   IF #Startup THEN
       "StationA".Access.Policy.Required[11] := 3;
       "StationB".Access.Policy.Required[11] := 3;
   END_IF;
   IF #Startup THEN
       IF NOT "FRK_AccessStorage".UsersCommissioned AND "FRK_LocalUsers".SchemaVersion = 0 AND "FRK_LocalUsers".Generation = 0 AND "FRK_LocalUsers".Checksum = DWORD#0 THEN
           "F_AccessBenchProvision"();
       END_IF;
       "StationA".Access.Policy.Required[2] := 1;
       "StationA".Access.Policy.Required[4] := 1;
       "StationA".Access.Policy.Required[5] := 1;
       "StationA".Access.Policy.Required[8] := 4;
       "StationA".Access.Policy.SessionTimeout := T#0ms;
       "StationB".Access.Policy.Required[2] := 1;
       "StationB".Access.Policy.Required[4] := 1;
       "StationB".Access.Policy.Required[5] := 1;
       "StationB".Access.Policy.Required[8] := 4;
       "StationB".Access.Policy.SessionTimeout := T#0ms;
       "GDB_AccessTest".HashData[0] := BYTE#16#00;
       "GDB_AccessTest".HashData[1] := BYTE#16#01;
       "GDB_AccessTest".HashData[2] := BYTE#16#02;
       "GDB_AccessTest".HashData[3] := BYTE#16#03;
       "GDB_AccessTest".HashData[4] := BYTE#16#04;
       "GDB_AccessTest".HashData[5] := BYTE#16#05;
       "GDB_AccessTest".HashData[6] := BYTE#16#06;
       "GDB_AccessTest".HashData[7] := BYTE#16#07;
       "GDB_AccessTest".HashData[8] := BYTE#16#08;
       "GDB_AccessTest".HashData[9] := BYTE#16#09;
       "GDB_AccessTest".HashData[10] := BYTE#16#0A;
       "GDB_AccessTest".HashData[11] := BYTE#16#0B;
       "GDB_AccessTest".HashData[12] := BYTE#16#0C;
       "GDB_AccessTest".HashData[13] := BYTE#16#0D;
       "GDB_AccessTest".HashData[14] := BYTE#16#0E;
       "GDB_AccessTest".HashData[15] := BYTE#16#0F;
       "GDB_AccessTest".HashData[16] := BYTE#16#10;
       "GDB_AccessTest".HashData[17] := BYTE#16#11;
       "GDB_AccessTest".HashData[18] := BYTE#16#12;
       "GDB_AccessTest".HashData[19] := BYTE#16#13;
       "GDB_AccessTest".HashData[20] := BYTE#16#14;
       "GDB_AccessTest".HashData[21] := BYTE#16#15;
       "GDB_AccessTest".HashData[22] := BYTE#16#16;
       "GDB_AccessTest".HashData[23] := BYTE#16#17;
       "GDB_AccessTest".HashData[24] := BYTE#16#18;
       "GDB_AccessTest".HashData[25] := BYTE#16#19;
       "GDB_AccessTest".HashData[26] := BYTE#16#1A;
       "GDB_AccessTest".HashData[27] := BYTE#16#1B;
       "GDB_AccessTest".HashData[28] := BYTE#16#1C;
       "GDB_AccessTest".HashData[29] := BYTE#16#1D;
       "GDB_AccessTest".HashData[30] := BYTE#16#1E;
       "GDB_AccessTest".HashData[31] := BYTE#16#1F;
       "GDB_AccessTest".HashData[32] := BYTE#16#20;
       "GDB_AccessTest".HashData[33] := BYTE#16#21;
       "GDB_AccessTest".HashData[34] := BYTE#16#22;
       "GDB_AccessTest".HashData[35] := BYTE#16#23;
       "GDB_AccessTest".HashData[36] := BYTE#16#24;
       "GDB_AccessTest".HashData[37] := BYTE#16#25;
       "GDB_AccessTest".HashData[38] := BYTE#16#26;
       "GDB_AccessTest".HashData[39] := BYTE#16#27;
       "GDB_AccessTest".HashData[40] := BYTE#16#28;
       "GDB_AccessTest".HashData[41] := BYTE#16#29;
       "GDB_AccessTest".HashData[42] := BYTE#16#2A;
       "GDB_AccessTest".HashData[43] := BYTE#16#2B;
       "GDB_AccessTest".HashData[44] := BYTE#16#2C;
       "GDB_AccessTest".HashData[45] := BYTE#16#2D;
       "GDB_AccessTest".HashData[46] := BYTE#16#2E;
       "GDB_AccessTest".HashData[47] := BYTE#16#2F;
       "GDB_AccessTest".HashOk := "FRK_Sha256Pin"(Data := "GDB_AccessTest".HashData, Size := 0, Digest := "GDB_AccessTest".Hash0);
       "GDB_AccessTest".HashData[0] := BYTE#16#61;
       "GDB_AccessTest".HashData[1] := BYTE#16#62;
       "GDB_AccessTest".HashData[2] := BYTE#16#63;
       "GDB_AccessTest".HashData[3] := BYTE#16#00;
       "GDB_AccessTest".HashData[4] := BYTE#16#00;
       "GDB_AccessTest".HashData[5] := BYTE#16#00;
       "GDB_AccessTest".HashData[6] := BYTE#16#00;
       "GDB_AccessTest".HashData[7] := BYTE#16#00;
       "GDB_AccessTest".HashData[8] := BYTE#16#00;
       "GDB_AccessTest".HashData[9] := BYTE#16#00;
       "GDB_AccessTest".HashData[10] := BYTE#16#00;
       "GDB_AccessTest".HashData[11] := BYTE#16#00;
       "GDB_AccessTest".HashData[12] := BYTE#16#00;
       "GDB_AccessTest".HashData[13] := BYTE#16#00;
       "GDB_AccessTest".HashData[14] := BYTE#16#00;
       "GDB_AccessTest".HashData[15] := BYTE#16#00;
       "GDB_AccessTest".HashData[16] := BYTE#16#00;
       "GDB_AccessTest".HashData[17] := BYTE#16#00;
       "GDB_AccessTest".HashData[18] := BYTE#16#00;
       "GDB_AccessTest".HashData[19] := BYTE#16#00;
       "GDB_AccessTest".HashData[20] := BYTE#16#00;
       "GDB_AccessTest".HashData[21] := BYTE#16#00;
       "GDB_AccessTest".HashData[22] := BYTE#16#00;
       "GDB_AccessTest".HashData[23] := BYTE#16#00;
       "GDB_AccessTest".HashData[24] := BYTE#16#00;
       "GDB_AccessTest".HashData[25] := BYTE#16#00;
       "GDB_AccessTest".HashData[26] := BYTE#16#00;
       "GDB_AccessTest".HashData[27] := BYTE#16#00;
       "GDB_AccessTest".HashData[28] := BYTE#16#00;
       "GDB_AccessTest".HashData[29] := BYTE#16#00;
       "GDB_AccessTest".HashData[30] := BYTE#16#00;
       "GDB_AccessTest".HashData[31] := BYTE#16#00;
       "GDB_AccessTest".HashData[32] := BYTE#16#00;
       "GDB_AccessTest".HashData[33] := BYTE#16#00;
       "GDB_AccessTest".HashData[34] := BYTE#16#00;
       "GDB_AccessTest".HashData[35] := BYTE#16#00;
       "GDB_AccessTest".HashData[36] := BYTE#16#00;
       "GDB_AccessTest".HashData[37] := BYTE#16#00;
       "GDB_AccessTest".HashData[38] := BYTE#16#00;
       "GDB_AccessTest".HashData[39] := BYTE#16#00;
       "GDB_AccessTest".HashData[40] := BYTE#16#00;
       "GDB_AccessTest".HashData[41] := BYTE#16#00;
       "GDB_AccessTest".HashData[42] := BYTE#16#00;
       "GDB_AccessTest".HashData[43] := BYTE#16#00;
       "GDB_AccessTest".HashData[44] := BYTE#16#00;
       "GDB_AccessTest".HashData[45] := BYTE#16#00;
       "GDB_AccessTest".HashData[46] := BYTE#16#00;
       "GDB_AccessTest".HashData[47] := BYTE#16#00;
       "GDB_AccessTest".HashOk := "FRK_Sha256Pin"(Data := "GDB_AccessTest".HashData, Size := 3, Digest := "GDB_AccessTest".Hash1);
       "GDB_AccessTest".HashData[0] := BYTE#16#00;
       "GDB_AccessTest".HashData[1] := BYTE#16#01;
       "GDB_AccessTest".HashData[2] := BYTE#16#02;
       "GDB_AccessTest".HashData[3] := BYTE#16#03;
       "GDB_AccessTest".HashData[4] := BYTE#16#04;
       "GDB_AccessTest".HashData[5] := BYTE#16#05;
       "GDB_AccessTest".HashData[6] := BYTE#16#06;
       "GDB_AccessTest".HashData[7] := BYTE#16#07;
       "GDB_AccessTest".HashData[8] := BYTE#16#08;
       "GDB_AccessTest".HashData[9] := BYTE#16#09;
       "GDB_AccessTest".HashData[10] := BYTE#16#0A;
       "GDB_AccessTest".HashData[11] := BYTE#16#0B;
       "GDB_AccessTest".HashData[12] := BYTE#16#0C;
       "GDB_AccessTest".HashData[13] := BYTE#16#0D;
       "GDB_AccessTest".HashData[14] := BYTE#16#0E;
       "GDB_AccessTest".HashData[15] := BYTE#16#0F;
       "GDB_AccessTest".HashData[16] := BYTE#16#10;
       "GDB_AccessTest".HashData[17] := BYTE#16#11;
       "GDB_AccessTest".HashData[18] := BYTE#16#12;
       "GDB_AccessTest".HashData[19] := BYTE#16#13;
       "GDB_AccessTest".HashData[20] := BYTE#16#14;
       "GDB_AccessTest".HashData[21] := BYTE#16#15;
       "GDB_AccessTest".HashData[22] := BYTE#16#16;
       "GDB_AccessTest".HashData[23] := BYTE#16#17;
       "GDB_AccessTest".HashData[24] := BYTE#16#18;
       "GDB_AccessTest".HashData[25] := BYTE#16#19;
       "GDB_AccessTest".HashData[26] := BYTE#16#1A;
       "GDB_AccessTest".HashData[27] := BYTE#16#1B;
       "GDB_AccessTest".HashData[28] := BYTE#16#1C;
       "GDB_AccessTest".HashData[29] := BYTE#16#1D;
       "GDB_AccessTest".HashData[30] := BYTE#16#1E;
       "GDB_AccessTest".HashData[31] := BYTE#16#1F;
       "GDB_AccessTest".HashData[32] := BYTE#16#20;
       "GDB_AccessTest".HashData[33] := BYTE#16#21;
       "GDB_AccessTest".HashData[34] := BYTE#16#22;
       "GDB_AccessTest".HashData[35] := BYTE#16#23;
       "GDB_AccessTest".HashData[36] := BYTE#16#24;
       "GDB_AccessTest".HashData[37] := BYTE#16#25;
       "GDB_AccessTest".HashData[38] := BYTE#16#26;
       "GDB_AccessTest".HashData[39] := BYTE#16#27;
       "GDB_AccessTest".HashData[40] := BYTE#16#28;
       "GDB_AccessTest".HashData[41] := BYTE#16#29;
       "GDB_AccessTest".HashData[42] := BYTE#16#2A;
       "GDB_AccessTest".HashData[43] := BYTE#16#2B;
       "GDB_AccessTest".HashData[44] := BYTE#16#2C;
       "GDB_AccessTest".HashData[45] := BYTE#16#2D;
       "GDB_AccessTest".HashData[46] := BYTE#16#2E;
       "GDB_AccessTest".HashData[47] := BYTE#16#2F;
       "GDB_AccessTest".HashOk := "FRK_Sha256Pin"(Data := "GDB_AccessTest".HashData, Size := 32, Digest := "GDB_AccessTest".Hash2);
       "GDB_AccessTest".HashData[0] := BYTE#16#00;
       "GDB_AccessTest".HashData[1] := BYTE#16#01;
       "GDB_AccessTest".HashData[2] := BYTE#16#02;
       "GDB_AccessTest".HashData[3] := BYTE#16#03;
       "GDB_AccessTest".HashData[4] := BYTE#16#04;
       "GDB_AccessTest".HashData[5] := BYTE#16#05;
       "GDB_AccessTest".HashData[6] := BYTE#16#06;
       "GDB_AccessTest".HashData[7] := BYTE#16#07;
       "GDB_AccessTest".HashData[8] := BYTE#16#08;
       "GDB_AccessTest".HashData[9] := BYTE#16#09;
       "GDB_AccessTest".HashData[10] := BYTE#16#0A;
       "GDB_AccessTest".HashData[11] := BYTE#16#0B;
       "GDB_AccessTest".HashData[12] := BYTE#16#0C;
       "GDB_AccessTest".HashData[13] := BYTE#16#0D;
       "GDB_AccessTest".HashData[14] := BYTE#16#0E;
       "GDB_AccessTest".HashData[15] := BYTE#16#0F;
       "GDB_AccessTest".HashData[16] := BYTE#16#10;
       "GDB_AccessTest".HashData[17] := BYTE#16#11;
       "GDB_AccessTest".HashData[18] := BYTE#16#12;
       "GDB_AccessTest".HashData[19] := BYTE#16#13;
       "GDB_AccessTest".HashData[20] := BYTE#16#14;
       "GDB_AccessTest".HashData[21] := BYTE#16#15;
       "GDB_AccessTest".HashData[22] := BYTE#16#16;
       "GDB_AccessTest".HashData[23] := BYTE#16#17;
       "GDB_AccessTest".HashData[24] := BYTE#16#18;
       "GDB_AccessTest".HashData[25] := BYTE#16#19;
       "GDB_AccessTest".HashData[26] := BYTE#16#1A;
       "GDB_AccessTest".HashData[27] := BYTE#16#1B;
       "GDB_AccessTest".HashData[28] := BYTE#16#1C;
       "GDB_AccessTest".HashData[29] := BYTE#16#1D;
       "GDB_AccessTest".HashData[30] := BYTE#16#1E;
       "GDB_AccessTest".HashData[31] := BYTE#16#1F;
       "GDB_AccessTest".HashData[32] := BYTE#16#20;
       "GDB_AccessTest".HashData[33] := BYTE#16#21;
       "GDB_AccessTest".HashData[34] := BYTE#16#22;
       "GDB_AccessTest".HashData[35] := BYTE#16#23;
       "GDB_AccessTest".HashData[36] := BYTE#16#24;
       "GDB_AccessTest".HashData[37] := BYTE#16#25;
       "GDB_AccessTest".HashData[38] := BYTE#16#26;
       "GDB_AccessTest".HashData[39] := BYTE#16#27;
       "GDB_AccessTest".HashData[40] := BYTE#16#28;
       "GDB_AccessTest".HashData[41] := BYTE#16#29;
       "GDB_AccessTest".HashData[42] := BYTE#16#2A;
       "GDB_AccessTest".HashData[43] := BYTE#16#2B;
       "GDB_AccessTest".HashData[44] := BYTE#16#2C;
       "GDB_AccessTest".HashData[45] := BYTE#16#2D;
       "GDB_AccessTest".HashData[46] := BYTE#16#2E;
       "GDB_AccessTest".HashData[47] := BYTE#16#2F;
       "GDB_AccessTest".HashOk := "FRK_Sha256Pin"(Data := "GDB_AccessTest".HashData, Size := 48, Digest := "GDB_AccessTest".Hash3);
       "GDB_RoutingTest".PermitOne := TRUE;
       "GDB_RoutingTest".PermitTwo := TRUE;
       "GDB_RoutingTest".RootManualPermit := TRUE;
       "GDB_RoutingTest".NestedFinish := FALSE;
       "GDB_RoutingTest".InnerFinish := FALSE;
       "GDB_RoutingTest".NestedAccessLock := FALSE;
       #ResultCode := RD_SYS_T(OUT => #StartupStamp);
       IF #ResultCode = 0 THEN
           "GDB_UnitTest".BootStamp := DTL_TO_LDT(#StartupStamp);
       END_IF;
       "GDB_UnitTest".Restarts := "GDB_UnitTest".Restarts + 1;
       "GDB_UnitTest".FinishCycle := FALSE;
       "GDB_UnitTest".Permit := TRUE;
       "GDB_UnitTest".FaultRoot := FALSE;
       "GDB_UnitTest".ExitHold := FALSE;
       "GDB_UnitTest".IssueChild := FALSE;
       "GDB_UnitTest".LockStart := FALSE;
       "GDB_UnitTest".ChildCommand := 2;
       "GDB_UnitTest".Verdict := 1;
       "GDB_UnitTest".Reason := 2003;
       "GDB_UnitTest".CarrierControl := 0;
       "FRK_UnitSetLocalCarrier"(Unit := "StationA".Unit,
                                 Index := 1);
   END_IF;
   "GDB_FraktalHal".Data.StationA.Cell.Clamp.Finish := "GDB_UnitTest".FinishCycle;
   "GDB_FraktalHal".Data.StationA.Cell.Clamp.Permit := "GDB_UnitTest".Permit;
   "GDB_FraktalHal".Data.StationA.Cell.Clamp.ExitHold := "GDB_UnitTest".ExitHold;
   "GDB_FraktalHal".Data.StationA.Cell.Clamp.BackgroundFault := "GDB_UnitTest".FaultRoot;
   "GDB_FraktalHal".Data.StationA.Cell.Clamp.Verdict := "GDB_UnitTest".Verdict;
   "GDB_FraktalHal".Data.StationA.Cell.Clamp.Diag.ReasonCode := "GDB_UnitTest".Reason;
   "GDB_FraktalHal".Data.StationA.Cell.Clamp.Diag.Description := WSTRING#'test.start.permit';
   "GDB_FraktalHal".Data.StationA.Cell.Clamp.Diag.SourcePath := WSTRING#'StationA.Cell.Clamp';
   IF "GDB_UnitTest".IssueChild THEN
       "StationA".Cell.Clamp.Command := "GDB_UnitTest".ChildCommand;
       "StationA".Cell.Clamp.Execute := TRUE;
       "GDB_UnitTest".IssueChild := FALSE;
   END_IF;
   CASE "GDB_UnitTest".CarrierControl OF
       1:
           "FRK_UnitSetLocalCarrier"(Unit := "StationA".Unit,
                                     Index := 1);
       2:
           "FRK_Carriers".Slots[1].Enabled := FALSE;
       3:
           "FRK_Carriers".Slots[1].Context.Uid := 'other';
       ELSE
           "GDB_UnitTest".CarrierControl := 0;
   END_CASE;
   "GDB_UnitTest".CarrierControl := 0;
   "GDB_FraktalHal".Data.StationA.Cell.Gate.Permit := "GDB_RoutingTest".PermitOne;
   IF "GDB_RoutingTest".PermitTwo THEN
       "GDB_FraktalHal".Data.StationA.Cell.Gate.Sample := 0;
   ELSE
       "GDB_FraktalHal".Data.StationA.Cell.Gate.Sample := 1;
   END_IF;
   "GDB_FraktalHal".Data.StationA.Cell.Gate.Diag.ReasonCode := 2002;
   "GDB_FraktalHal".Data.StationA.Cell.Gate.Diag.Description := WSTRING#'test.manual.first';
   "GDB_FraktalHal".Data.StationA.Cell.Gate.LaterDiag.ReasonCode := 2003;
   "GDB_FraktalHal".Data.StationA.Cell.Gate.LaterDiag.Description := WSTRING#'test.manual.second';
   "GDB_FraktalHal".Data.StationA.Satellite.Cell.Clamp.Permit := "GDB_RoutingTest".RootManualPermit;
   "GDB_FraktalHal".Data.StationA.Satellite.Cell.Clamp.Diag.SourcePath := WSTRING#'StationA.Satellite.Cell.Clamp';
   "GDB_FraktalHal".Data.StationA.Satellite.Cell.Clamp.Diag.Description := WSTRING#'test.nested.permit';
   "GDB_FraktalHal".Data.StationA.Satellite.Cell.Clamp.Diag.ReasonCode := 2002;
   "GDB_FraktalHal".Data.StationA.Satellite.Inner.Cell.Clamp.Permit := TRUE;
   "GDB_FraktalHal".Data.StationA.Satellite.Cell.Clamp.Finish := "GDB_RoutingTest".NestedFinish;
   "GDB_FraktalHal".Data.StationA.Satellite.Inner.Cell.Clamp.Finish := "GDB_RoutingTest".InnerFinish;
   IF "GDB_RoutingTest".NestedAccessLock THEN
       "StationA".Satellite.Access.Policy.Required[5] := 4;
   ELSE
       "StationA".Satellite.Access.Policy.Required[5] := 0;
   END_IF;
   IF "GDB_RoutingTest".LocalPulse THEN
       "GDB_RoutingTest".LocalRequest.Kind := "GDB_RoutingTest".LocalKind;
       "GDB_RoutingTest".LocalRequest.IntValue := "GDB_RoutingTest".LocalValue;
       "FRK_UnitOperation"(Core := "StationA".Satellite.Core,
                           Unit := "StationA".Satellite.Unit,
                           Status := "StationA".Satellite.Status,
                           Policy := "StationA".Satellite.ModePolicy,
                           Access := "StationA".Satellite.Access,
                           Supported := "StationA".Satellite.SupportedModesPublished,
                           Request := "GDB_RoutingTest".LocalRequest,
                           Response := "FRK_UnitScratch".Response,
                           Trusted := FALSE);
       "GDB_RoutingTest".LocalAccepted := "FRK_UnitScratch".Response.Accepted;
       "GDB_RoutingTest".LocalFirstKind := -1;
       IF "FRK_UnitScratch".Response.Report.Count > 0 THEN
           "GDB_RoutingTest".LocalFirstKind := "FRK_UnitScratch".Response.Report.Reasons[1].Kind;
       END_IF;
       "GDB_RoutingTest".LocalPulse := FALSE;
   END_IF;
   "StationA".Access.ProviderEnabled := NOT "GDB_AccessTest".ProviderOff;
   "StationB".Access.ProviderEnabled := NOT "GDB_AccessTest".ProviderOff;
   "StationA".AlarmLog.SinkEnabled := TRUE;
   "StationB".AlarmLog.SinkEnabled := TRUE;
   "GDB_FraktalHal".Data.StationA.Cell.Clamp.Sample := "GDB_StateAlarmTest".Position;
   IF "GDB_StateAlarmTest".ClearLog THEN
       "FRK_AlarmBegin"(AlarmLog := "StationA".AlarmLog,
                        Startup := TRUE);
       "GDB_StateAlarmTest".SinkCome := 0;
       "GDB_StateAlarmTest".SinkClose := 0;
       "GDB_StateAlarmTest".ClearLog := FALSE;
   END_IF;
   IF "GDB_StateAlarmTest".RaisePulse THEN
       "GDB_StateAlarmTest".Slot := "FRK_AlarmRaise"(AlarmLog := "StationA".AlarmLog, Diag := "GDB_StateAlarmTest".Diag, ResetClass := "GDB_StateAlarmTest".ResetClass);
       "GDB_StateAlarmTest".RaisePulse := FALSE;
   END_IF;
   IF "GDB_StateAlarmTest".GonePulse THEN
       "GDB_StateAlarmTest".GoneAccepted := "FRK_AlarmGone"(AlarmLog := "StationA".AlarmLog, Slot := "GDB_StateAlarmTest".Slot);
       "GDB_StateAlarmTest".GonePulse := FALSE;
   END_IF;
   IF "GDB_StateAlarmTest".FillPulse THEN
       FOR #SlotIndex := 1 TO "GDB_StateAlarmTest".FillCount DO
           #Taken := "FRK_AlarmRaise"(AlarmLog := "StationA".AlarmLog, Diag := "GDB_StateAlarmTest".Diag, ResetClass := "GDB_StateAlarmTest".ResetClass);
           IF "GDB_StateAlarmTest".ResetClass = 0 THEN
               #Accepted := "FRK_AlarmGone"(AlarmLog := "StationA".AlarmLog, Slot := #Taken);
           END_IF;
       END_FOR;
       "GDB_StateAlarmTest".FillPulse := FALSE;
   END_IF;
   IF "GDB_StateAlarmTest".CauseLive THEN
       IF "GDB_StateAlarmTest".CauseSlot = 0 THEN
           "GDB_StateAlarmTest".CauseSlot := "FRK_AlarmRaise"(AlarmLog := "StationA".AlarmLog, Diag := "GDB_StateAlarmTest".Diag, ResetClass := 1);
       ELSIF "StationA".AlarmLog.Active["GDB_StateAlarmTest".CauseSlot].State = 0 THEN
           "GDB_StateAlarmTest".CauseSlot := "FRK_AlarmRaise"(AlarmLog := "StationA".AlarmLog, Diag := "GDB_StateAlarmTest".Diag, ResetClass := 1);
       END_IF;
   ELSIF "GDB_StateAlarmTest".CauseSlot > 0 THEN
       #Accepted := "FRK_AlarmGone"(AlarmLog := "StationA".AlarmLog, Slot := "GDB_StateAlarmTest".CauseSlot);
       "GDB_StateAlarmTest".CauseSlot := 0;
   END_IF;
   "FRK_StateSweep"(Flags := "GDB_StateAlarmTest".StandaloneFlags,
                    Count := "GDB_StateAlarmTest".StandaloneCount,
                    Touched := "GDB_StateAlarmTest".Touched,
                    Startup := #Startup);
   IF "GDB_StateAlarmTest".PublishState THEN
       "GDB_StateAlarmTest".StandaloneReturn := "FRK_State"(Idx := "GDB_StateAlarmTest".StateIndex, Key := 'project.state.atHome', Ok := "GDB_StateAlarmTest".StateValue, Flags := "GDB_StateAlarmTest".StandaloneFlags, Count := "GDB_StateAlarmTest".StandaloneCount, Touched := "GDB_StateAlarmTest".Touched);
   END_IF;
   "FRK_ConfigRuntime".Unavailable := "GDB_ConfigTest".Unavailable;
   IF "GDB_ConfigTest".BlockRestore THEN
       "StationA".ConfigPersist.RestorePolicy := 1;
   ELSE
       "StationA".ConfigPersist.RestorePolicy := 0;
   END_IF;
   IF "GDB_ConfigTest".CorruptPulse THEN
       "GDB_ConfigTest".CorruptSlot := "FRK_ConfigFind"(Scope := "GDB_ConfigTest".CorruptScope, Key := "GDB_ConfigTest".CorruptKey, ModelCode := "GDB_ConfigTest".CorruptModel);
       IF "GDB_ConfigTest".CorruptSlot > 0 THEN
           "FRK_ConfigStore".Rows["GDB_ConfigTest".CorruptSlot].SchemaVersion := "GDB_ConfigTest".CorruptSchema;
           "FRK_ConfigStore".Rows["GDB_ConfigTest".CorruptSlot].Record.ValueText := "GDB_ConfigTest".CorruptText;
       END_IF;
       "GDB_ConfigTest".CorruptPulse := FALSE;
   END_IF;
END_FUNCTION

FUNCTION "F_ConfigSetBench" : Void   // FC173, SCL
{ S7_Optimized_Access := 'TRUE' }
VERSION : 0.1
// Test-only tampering: the production retained store stays inaccessible.
// stored: AutoNumber true, IsIECCheckEnabled false, SetENOAutomatically false, UDAEnableTagReadback false
   VAR_TEMP
      Slot : Int;
      Index : Int;
   END_VAR
BEGIN

   IF NOT "GDB_ConfigSetTest".Corrupt THEN
       RETURN;
   END_IF;
   "GDB_ConfigSetTest".Corrupt := FALSE;
   #Slot := "FRK_SetFind"(RootIndex := 1, SetName := "GDB_ConfigSetTest".SetName);
   "GDB_ConfigSetTest".Slot := #Slot;
   IF #Slot = 0 THEN
       RETURN;
   END_IF;
   #Index := "FRK_SetStore".Sets[1, #Slot].Info.RecordCount;
   "GDB_ConfigSetTest".RecordScope := "FRK_SetStore".Sets[1, #Slot].Records[#Index].Scope;
   "GDB_ConfigSetTest".RecordKey := "FRK_SetStore".Sets[1, #Slot].Records[#Index].WriteKey;
   CASE "GDB_ConfigSetTest".Field OF
       1:
           "FRK_SetStore".Sets[1, #Slot].Records[#Index].ValueText := "GDB_ConfigSetTest".Text;
       2:
           "FRK_SetStore".Sets[1, #Slot].Records[#Index].Revision := 99;
       3:
           "FRK_SetStore".Sets[1, #Slot].Records[#Index].ValueType := 99;
       4:
           "FRK_SetStore".Sets[1, #Slot].Records[#Index].WriteKey := 'unknown';
       5:
           "FRK_SetStore".Sets[1, #Slot].Records[#Index].Scope := 'StationB';
       6:
           "FRK_SetStore".Sets[1, #Slot].Info.RecordCount := #Index - 1;
       7:
           "FRK_SetStore".Sets[1, #Slot].Records[#Index] := "FRK_SetStore".Sets[1, #Slot].Records[1];
       ELSE
           RETURN;
   END_CASE;
END_FUNCTION

FUNCTION "F_DecisionBench" : Void   // FC172, SCL
{ S7_Optimized_Access := 'TRUE' }
VERSION : 0.1
// stored: AutoNumber true, IsIECCheckEnabled false, SetENOAutomatically false, UDAEnableTagReadback false
   VAR_TEMP
      Root : DInt;
      Peer : DInt;
      Nested : DInt;
      Slot : Int;
      CaseNo : Int;
      RootPath : WString[255];
      PeerPath : WString[255];
      NestedPath : WString[255];
      "A" : Bool;
      "B" : Bool;
      C : Bool;
      Ok : Bool;
      Answer : Int;
      Head : Int;
   END_VAR
BEGIN

   IF "GDB_DecisionTest".Done OR "FRK_Registry".Fault THEN
       RETURN;
   END_IF;
   #Root := "StationA".Core.RegIndex;
   #Peer := "StationB".Core.RegIndex;
   #Nested := "StationA".Satellite.Core.RegIndex;
   IF #Root <= 0 OR #Peer <= 0 OR #Nested <= 0 THEN
       RETURN;
   END_IF;
   #RootPath := STRING_TO_WSTRING("StationA".Status.Name);
   #PeerPath := STRING_TO_WSTRING("StationB".Status.Name);
   #NestedPath := STRING_TO_WSTRING("StationA".Satellite.Status.Name);
   #Slot := "FRK_DecisionRoot"(Owner := #Root, Create := TRUE);
   "GDB_DecisionTest".Total := 28;
   FOR #CaseNo := 1 TO 28 DO
       "FRK_DecisionCyclic"(Owner := #Root,
                            Busy := FALSE,
                            Reset := TRUE,
                            AlarmLog := "GDB_DecisionTest".Log);
       "FRK_DecisionCyclic"(Owner := #Peer,
                            Busy := FALSE,
                            Reset := TRUE,
                            AlarmLog := "GDB_DecisionTest".Log);
       "GDB_DecisionTest".WorkRequest := "FRK_Decisions".EmptyRequest;
       "GDB_DecisionTest".WorkRequest.Prompt := WSTRING#'test.decision.prompt';
       "GDB_DecisionTest".WorkRequest.Options[1] := 'test.decision.optionOne';
       "GDB_DecisionTest".WorkRequest.Options[2] := 'test.decision.optionTwo';
       "GDB_DecisionTest".WorkHmiRequest := "GDB_DecisionTest".EmptyHmiRequest;
       "GDB_DecisionTest".WorkHmiResponse := "GDB_DecisionTest".EmptyHmiResponse;
       "GDB_DecisionTest".WorkReport := "GDB_DecisionTest".EmptyReport;
       "GDB_DecisionTest".WorkPublished := "FRK_Decisions".EmptyRequest;
       "GDB_DecisionTest".WorkReport.Count := 0;
       "GDB_DecisionTest".WorkReport.Released := TRUE;
       #Ok := FALSE;
       CASE #CaseNo OF
           1: // invalid_owner
               #A := "FRK_DecisionAsk"(Owner := 0, OwnerPath := #RootPath, Request := "GDB_DecisionTest".WorkRequest, AlarmLog := "GDB_DecisionTest".Log);
               #Ok := NOT #A;
           2: // root_publication
               #A := "FRK_DecisionAsk"(Owner := #Root, OwnerPath := #RootPath, Request := "GDB_DecisionTest".WorkRequest, AlarmLog := "GDB_DecisionTest".Log);
               "FRK_DecisionPublish"(Owner := #Root,
                                     Decision := "GDB_DecisionTest".WorkPublished,
                                     DecisionAnswer := #Answer);
               #Ok := #A AND "GDB_DecisionTest".WorkPublished.Prompt = "GDB_DecisionTest".WorkRequest.Prompt AND "GDB_DecisionTest".WorkPublished.SourcePath = #RootPath AND #Answer = 0;
           3: // idempotent_no_flood
               #A := "FRK_DecisionAsk"(Owner := #Root, OwnerPath := #RootPath, Request := "GDB_DecisionTest".WorkRequest, AlarmLog := "GDB_DecisionTest".Log);
               #Head := "GDB_DecisionTest".Log.RingHead;
               #A := "FRK_DecisionAsk"(Owner := #Root, OwnerPath := #RootPath, Request := "GDB_DecisionTest".WorkRequest, AlarmLog := "GDB_DecisionTest".Log);
               #Ok := #A AND #Head = "GDB_DecisionTest".Log.RingHead;
           4: // overlap_preserves_first
               #A := "FRK_DecisionAsk"(Owner := #Root, OwnerPath := #RootPath, Request := "GDB_DecisionTest".WorkRequest, AlarmLog := "GDB_DecisionTest".Log);
               "GDB_DecisionTest".WorkRequest.Prompt := WSTRING#'test.decision.different';
               #A := "FRK_DecisionAsk"(Owner := #Root, OwnerPath := #RootPath, Request := "GDB_DecisionTest".WorkRequest, AlarmLog := "GDB_DecisionTest".Log);
               #Head := "GDB_DecisionTest".Log.RingHead;
               #B := #A;
               #A := "FRK_DecisionAsk"(Owner := #Root, OwnerPath := #RootPath, Request := "GDB_DecisionTest".WorkRequest, AlarmLog := "GDB_DecisionTest".Log);
               "FRK_DecisionPublish"(Owner := #Root,
                                     Decision := "GDB_DecisionTest".WorkPublished,
                                     DecisionAnswer := #Answer);
               #Ok := NOT #B AND NOT #A AND "GDB_DecisionTest".WorkPublished.Prompt = WSTRING#'test.decision.prompt' AND #Head = "GDB_DecisionTest".Log.RingHead;
           5: // nested_request_root_mirror
               #A := "FRK_DecisionAsk"(Owner := #Nested, OwnerPath := #NestedPath, Request := "GDB_DecisionTest".WorkRequest, AlarmLog := "GDB_DecisionTest".Log);
               "FRK_DecisionPublish"(Owner := #Root,
                                     Decision := "GDB_DecisionTest".WorkPublished,
                                     DecisionAnswer := #Answer);
               #B := "GDB_DecisionTest".WorkPublished.SourcePath = #NestedPath;
               "FRK_DecisionPublish"(Owner := #Nested,
                                     Decision := "GDB_DecisionTest".WorkPublished,
                                     DecisionAnswer := #Answer);
               #Ok := #A AND #B AND "GDB_DecisionTest".WorkPublished.Prompt = WSTRING#'';
           6: // peer_roots_independent
               #A := "FRK_DecisionAsk"(Owner := #Root, OwnerPath := #RootPath, Request := "GDB_DecisionTest".WorkRequest, AlarmLog := "GDB_DecisionTest".Log);
               "GDB_DecisionTest".WorkRequest.Prompt := WSTRING#'test.decision.peer';
               #B := "FRK_DecisionAsk"(Owner := #Peer, OwnerPath := #PeerPath, Request := "GDB_DecisionTest".WorkRequest, AlarmLog := "GDB_DecisionTest".Log);
               "FRK_DecisionPublish"(Owner := #Root,
                                     Decision := "GDB_DecisionTest".WorkPublished,
                                     DecisionAnswer := #Answer);
               #Ok := #A AND #B AND "GDB_DecisionTest".WorkPublished.Prompt = WSTRING#'test.decision.prompt';
               "FRK_DecisionPublish"(Owner := #Peer,
                                     Decision := "GDB_DecisionTest".WorkPublished,
                                     DecisionAnswer := #Answer);
               #Ok := #Ok AND "GDB_DecisionTest".WorkPublished.Prompt = WSTRING#'test.decision.peer';
           7: // zero_timeout_indefinite
               #A := "FRK_DecisionAsk"(Owner := #Root, OwnerPath := #RootPath, Request := "GDB_DecisionTest".WorkRequest, AlarmLog := "GDB_DecisionTest".Log);
               "FRK_Decisions".Slots[#Slot].AskedAt := "FRK_Clock".NowMs - 5000;
               "FRK_DecisionCyclic"(Owner := #Root,
                                    Busy := TRUE,
                                    Reset := FALSE,
                                    AlarmLog := "GDB_DecisionTest".Log);
               "FRK_DecisionPublish"(Owner := #Root,
                                     Decision := "GDB_DecisionTest".WorkPublished,
                                     DecisionAnswer := #Answer);
               #Ok := #A AND #Answer = 0 AND "GDB_DecisionTest".WorkPublished.Prompt <> WSTRING#'';
           8: // finite_timeout_default
               "GDB_DecisionTest".WorkRequest.Timeout := T#2ms;
               "GDB_DecisionTest".WorkRequest.Default := 2;
               #A := "FRK_DecisionAsk"(Owner := #Root, OwnerPath := #RootPath, Request := "GDB_DecisionTest".WorkRequest, AlarmLog := "GDB_DecisionTest".Log);
               "FRK_Decisions".Slots[#Slot].AskedAt := "FRK_Clock".NowMs - 5;
               "FRK_DecisionCyclic"(Owner := #Root,
                                    Busy := TRUE,
                                    Reset := FALSE,
                                    AlarmLog := "GDB_DecisionTest".Log);
               #Answer := "FRK_DecisionTake"(Owner := #Root, AlarmLog := "GDB_DecisionTest".Log);
               #Ok := #A AND #Answer = 2;
           9: // finite_requires_default
               "GDB_DecisionTest".WorkRequest.Timeout := T#2ms;
               #A := "FRK_DecisionAsk"(Owner := #Root, OwnerPath := #RootPath, Request := "GDB_DecisionTest".WorkRequest, AlarmLog := "GDB_DecisionTest".Log);
               #Ok := NOT #A;
           10: // default_must_be_offered
               "GDB_DecisionTest".WorkRequest.Default := 3;
               #A := "FRK_DecisionAsk"(Owner := #Root, OwnerPath := #RootPath, Request := "GDB_DecisionTest".WorkRequest, AlarmLog := "GDB_DecisionTest".Log);
               #Ok := NOT #A;
           11: // negative_timeout_rejected
               "GDB_DecisionTest".WorkRequest.Timeout := T#-1ms;
               #A := "FRK_DecisionAsk"(Owner := #Root, OwnerPath := #RootPath, Request := "GDB_DecisionTest".WorkRequest, AlarmLog := "GDB_DecisionTest".Log);
               #Ok := NOT #A;
           12: // option_zero_rejected
               #A := "FRK_DecisionAsk"(Owner := #Root, OwnerPath := #RootPath, Request := "GDB_DecisionTest".WorkRequest, AlarmLog := "GDB_DecisionTest".Log);
               "GDB_DecisionTest".WorkReport.Released := TRUE;
               #B := "FRK_DecisionSubmit"(Owner := #Root, OwnerPath := #RootPath, Option := 0, Busy := TRUE, Permit := TRUE, Report := "GDB_DecisionTest".WorkReport);
               #Ok := #A AND NOT #B AND NOT "GDB_DecisionTest".WorkReport.Released;
           13: // unoffered_option_rejected
               #A := "FRK_DecisionAsk"(Owner := #Root, OwnerPath := #RootPath, Request := "GDB_DecisionTest".WorkRequest, AlarmLog := "GDB_DecisionTest".Log);
               "GDB_DecisionTest".WorkReport.Released := TRUE;
               #B := "FRK_DecisionSubmit"(Owner := #Root, OwnerPath := #RootPath, Option := 3, Busy := TRUE, Permit := TRUE, Report := "GDB_DecisionTest".WorkReport);
               #Ok := #A AND NOT #B AND NOT "GDB_DecisionTest".WorkReport.Released;
           14: // answer_consumed_once
               #A := "FRK_DecisionAsk"(Owner := #Root, OwnerPath := #RootPath, Request := "GDB_DecisionTest".WorkRequest, AlarmLog := "GDB_DecisionTest".Log);
               "GDB_DecisionTest".WorkReport.Released := TRUE;
               #B := "FRK_DecisionSubmit"(Owner := #Root, OwnerPath := #RootPath, Option := 1, Busy := TRUE, Permit := TRUE, Report := "GDB_DecisionTest".WorkReport);
               #Answer := "FRK_DecisionTake"(Owner := #Root, AlarmLog := "GDB_DecisionTest".Log);
               #Ok := #A AND #B AND #Answer = 1;
               #Answer := "FRK_DecisionTake"(Owner := #Root, AlarmLog := "GDB_DecisionTest".Log);
               #Ok := #Ok AND #Answer = 0;
           15: // duplicate_answer_rejected
               #A := "FRK_DecisionAsk"(Owner := #Root, OwnerPath := #RootPath, Request := "GDB_DecisionTest".WorkRequest, AlarmLog := "GDB_DecisionTest".Log);
               "GDB_DecisionTest".WorkReport.Released := TRUE;
               #B := "FRK_DecisionSubmit"(Owner := #Root, OwnerPath := #RootPath, Option := 1, Busy := TRUE, Permit := TRUE, Report := "GDB_DecisionTest".WorkReport);
               #C := #B;
               "GDB_DecisionTest".WorkReport.Released := TRUE;
               #B := "FRK_DecisionSubmit"(Owner := #Root, OwnerPath := #RootPath, Option := 2, Busy := TRUE, Permit := TRUE, Report := "GDB_DecisionTest".WorkReport);
               #Answer := "FRK_DecisionTake"(Owner := #Root, AlarmLog := "GDB_DecisionTest".Log);
               #Ok := #A AND #C AND NOT #B AND #Answer = 1;
           16: // interlock_denies_answer
               #A := "FRK_DecisionAsk"(Owner := #Root, OwnerPath := #RootPath, Request := "GDB_DecisionTest".WorkRequest, AlarmLog := "GDB_DecisionTest".Log);
               "GDB_DecisionTest".WorkReport.Released := TRUE;
               #B := "FRK_DecisionSubmit"(Owner := #Root, OwnerPath := #RootPath, Option := 1, Busy := TRUE, Permit := FALSE, Report := "GDB_DecisionTest".WorkReport);
               #Ok := #A AND NOT #B AND NOT "GDB_DecisionTest".WorkReport.Released AND "FRK_Decisions".Slots[#Slot].Answer = 0;
           17: // release_denial_preserved
               #A := "FRK_DecisionAsk"(Owner := #Root, OwnerPath := #RootPath, Request := "GDB_DecisionTest".WorkRequest, AlarmLog := "GDB_DecisionTest".Log);
               "GDB_DecisionTest".WorkReport.Released := FALSE;
               #B := "FRK_DecisionSubmit"(Owner := #Root, OwnerPath := #RootPath, Option := 1, Busy := TRUE, Permit := TRUE, Report := "GDB_DecisionTest".WorkReport);
               #Ok := #A AND NOT #B AND "FRK_Decisions".Slots[#Slot].Answer = 0;
           18: // reset_withdraws
               #A := "FRK_DecisionAsk"(Owner := #Root, OwnerPath := #RootPath, Request := "GDB_DecisionTest".WorkRequest, AlarmLog := "GDB_DecisionTest".Log);
               "FRK_DecisionCyclic"(Owner := #Root,
                                    Busy := TRUE,
                                    Reset := TRUE,
                                    AlarmLog := "GDB_DecisionTest".Log);
               #Ok := #A AND "FRK_Decisions".Slots[#Slot].Request.Prompt = WSTRING#'';
           19: // idle_fault_abort_withdraws
               #A := "FRK_DecisionAsk"(Owner := #Root, OwnerPath := #RootPath, Request := "GDB_DecisionTest".WorkRequest, AlarmLog := "GDB_DecisionTest".Log);
               "FRK_DecisionCyclic"(Owner := #Root,
                                    Busy := FALSE,
                                    Reset := FALSE,
                                    AlarmLog := "GDB_DecisionTest".Log);
               #Ok := #A AND "FRK_Decisions".Slots[#Slot].Request.Prompt = WSTRING#'';
           20: // nested_idle_cannot_cancel
               #A := "FRK_DecisionAsk"(Owner := #Root, OwnerPath := #RootPath, Request := "GDB_DecisionTest".WorkRequest, AlarmLog := "GDB_DecisionTest".Log);
               "FRK_DecisionCyclic"(Owner := #Nested,
                                    Busy := FALSE,
                                    Reset := TRUE,
                                    AlarmLog := "GDB_DecisionTest".Log);
               #Ok := #A AND "FRK_Decisions".Slots[#Slot].Request.Prompt <> WSTRING#'';
           21: // operator_wins_timeout_scan
               "GDB_DecisionTest".WorkRequest.Timeout := T#2ms;
               "GDB_DecisionTest".WorkRequest.Default := 2;
               #A := "FRK_DecisionAsk"(Owner := #Root, OwnerPath := #RootPath, Request := "GDB_DecisionTest".WorkRequest, AlarmLog := "GDB_DecisionTest".Log);
               "FRK_Decisions".Slots[#Slot].AskedAt := "FRK_Clock".NowMs - 5;
               "GDB_DecisionTest".WorkReport.Released := TRUE;
               #B := "FRK_DecisionSubmit"(Owner := #Root, OwnerPath := #RootPath, Option := 1, Busy := TRUE, Permit := TRUE, Report := "GDB_DecisionTest".WorkReport);
               "FRK_DecisionCyclic"(Owner := #Root,
                                    Busy := TRUE,
                                    Reset := FALSE,
                                    AlarmLog := "GDB_DecisionTest".Log);
               #Answer := "FRK_DecisionTake"(Owner := #Root, AlarmLog := "GDB_DecisionTest".Log);
               #Ok := #A AND #B AND #Answer = 1;
           22: // nested_mailbox_cannot_answer
               #A := "FRK_DecisionAsk"(Owner := #Root, OwnerPath := #RootPath, Request := "GDB_DecisionTest".WorkRequest, AlarmLog := "GDB_DecisionTest".Log);
               "GDB_DecisionTest".WorkReport.Released := TRUE;
               #B := "FRK_DecisionSubmit"(Owner := #Nested, OwnerPath := #NestedPath, Option := 1, Busy := TRUE, Permit := TRUE, Report := "GDB_DecisionTest".WorkReport);
               #Ok := #A AND NOT #B AND "FRK_Decisions".Slots[#Slot].Answer = 0;
           23: // audit_is_closed_nonblocking
               #A := "FRK_DecisionAsk"(Owner := #Root, OwnerPath := #RootPath, Request := "GDB_DecisionTest".WorkRequest, AlarmLog := "GDB_DecisionTest".Log);
               "GDB_DecisionTest".WorkReport.Released := TRUE;
               #B := "FRK_DecisionSubmit"(Owner := #Root, OwnerPath := #RootPath, Option := 1, Busy := TRUE, Permit := TRUE, Report := "GDB_DecisionTest".WorkReport);
               #Answer := "FRK_DecisionTake"(Owner := #Root, AlarmLog := "GDB_DecisionTest".Log);
               #Ok := #A AND #B AND #Answer = 1 AND NOT "GDB_DecisionTest".Log.Blocking AND "GDB_DecisionTest".Log.NActive = 0;
           24: // unit_access_gate
               #A := "FRK_DecisionAsk"(Owner := #Root, OwnerPath := #RootPath, Request := "GDB_DecisionTest".WorkRequest, AlarmLog := "GDB_DecisionTest".Log);
               "GDB_DecisionTest".WorkTestCore := "StationA".Core;
               "GDB_DecisionTest".WorkTestCore.Exec := 1;
               "GDB_DecisionTest".WorkTestUnit := "StationA".Unit;
               "GDB_DecisionTest".WorkTestUnit.Permit := TRUE;
               "GDB_DecisionTest".WorkTestAccess := "StationA".Access;
               "GDB_DecisionTest".WorkTestAccess.CurrentLevel := 0;
               "GDB_DecisionTest".WorkTestAccess.Policy.Required[5] := 1;
               "GDB_DecisionTest".WorkHmiRequest.Kind := 10;
               "GDB_DecisionTest".WorkHmiRequest.IntValue := 1;
               "FRK_UnitOperation"(Core := "GDB_DecisionTest".WorkTestCore,
                                   Unit := "GDB_DecisionTest".WorkTestUnit,
                                   Status := "StationA".Status,
                                   Policy := "StationA".ModePolicy,
                                   Access := "GDB_DecisionTest".WorkTestAccess,
                                   Response := "GDB_DecisionTest".WorkHmiResponse,
                                   Supported := "StationA".SupportedModesPublished,
                                   Request := "GDB_DecisionTest".WorkHmiRequest,
                                   Trusted := FALSE);
               #C := NOT "GDB_DecisionTest".WorkHmiResponse.Accepted AND NOT "GDB_DecisionTest".WorkHmiResponse.Report.Released AND "FRK_Decisions".Slots[#Slot].Answer = 0;
               "GDB_DecisionTest".WorkTestAccess.CurrentLevel := 1;
               "FRK_UnitOperation"(Core := "GDB_DecisionTest".WorkTestCore,
                                   Unit := "GDB_DecisionTest".WorkTestUnit,
                                   Status := "StationA".Status,
                                   Policy := "StationA".ModePolicy,
                                   Access := "GDB_DecisionTest".WorkTestAccess,
                                   Response := "GDB_DecisionTest".WorkHmiResponse,
                                   Supported := "StationA".SupportedModesPublished,
                                   Request := "GDB_DecisionTest".WorkHmiRequest,
                                   Trusted := FALSE);
               #Answer := "FRK_DecisionTake"(Owner := #Root, AlarmLog := "GDB_DecisionTest".Log);
               #Ok := #A AND #C AND "GDB_DecisionTest".WorkHmiResponse.Accepted AND #Answer = 1;
           25: // unit_idle_rejects_answer
               #A := "FRK_DecisionAsk"(Owner := #Root, OwnerPath := #RootPath, Request := "GDB_DecisionTest".WorkRequest, AlarmLog := "GDB_DecisionTest".Log);
               "GDB_DecisionTest".WorkTestCore := "StationA".Core;
               "GDB_DecisionTest".WorkTestCore.Exec := 0;
               "GDB_DecisionTest".WorkTestUnit := "StationA".Unit;
               "GDB_DecisionTest".WorkTestUnit.Permit := TRUE;
               "GDB_DecisionTest".WorkTestAccess := "StationA".Access;
               "GDB_DecisionTest".WorkTestAccess.CurrentLevel := 4;
               "GDB_DecisionTest".WorkHmiRequest.Kind := 10;
               "GDB_DecisionTest".WorkHmiRequest.IntValue := 1;
               "FRK_UnitOperation"(Core := "GDB_DecisionTest".WorkTestCore,
                                   Unit := "GDB_DecisionTest".WorkTestUnit,
                                   Status := "StationA".Status,
                                   Policy := "StationA".ModePolicy,
                                   Access := "GDB_DecisionTest".WorkTestAccess,
                                   Response := "GDB_DecisionTest".WorkHmiResponse,
                                   Supported := "StationA".SupportedModesPublished,
                                   Request := "GDB_DecisionTest".WorkHmiRequest,
                                   Trusted := FALSE);
               #Ok := #A AND NOT "GDB_DecisionTest".WorkHmiResponse.Accepted AND "FRK_Decisions".Slots[#Slot].Answer = 0;
           26: // forged_source_rejected
               "GDB_DecisionTest".WorkRequest.SourcePath := WSTRING#'OtherRoot';
               #A := "FRK_DecisionAsk"(Owner := #Root, OwnerPath := #RootPath, Request := "GDB_DecisionTest".WorkRequest, AlarmLog := "GDB_DecisionTest".Log);
               #Ok := NOT #A;
           27: // only_raiser_consumes
               #A := "FRK_DecisionAsk"(Owner := #Root, OwnerPath := #RootPath, Request := "GDB_DecisionTest".WorkRequest, AlarmLog := "GDB_DecisionTest".Log);
               "GDB_DecisionTest".WorkReport.Released := TRUE;
               #B := "FRK_DecisionSubmit"(Owner := #Root, OwnerPath := #RootPath, Option := 1, Busy := TRUE, Permit := TRUE, Report := "GDB_DecisionTest".WorkReport);
               #Answer := "FRK_DecisionTake"(Owner := #Nested, AlarmLog := "GDB_DecisionTest".Log);
               #C := #Answer = 0;
               #Answer := "FRK_DecisionTake"(Owner := #Root, AlarmLog := "GDB_DecisionTest".Log);
               #Ok := #A AND #B AND #C AND #Answer = 1;
           28: // root_withdraws_nested_request
               #A := "FRK_DecisionAsk"(Owner := #Nested, OwnerPath := #NestedPath, Request := "GDB_DecisionTest".WorkRequest, AlarmLog := "GDB_DecisionTest".Log);
               "FRK_DecisionCyclic"(Owner := #Root,
                                    Busy := FALSE,
                                    Reset := FALSE,
                                    AlarmLog := "GDB_DecisionTest".Log);
               #Ok := #A AND "FRK_Decisions".Slots[#Slot].Request.Prompt = WSTRING#'';
       END_CASE;
       "GDB_DecisionTest".Checks[#CaseNo] := #Ok;
       IF #Ok THEN
           "GDB_DecisionTest".Passed := "GDB_DecisionTest".Passed + 1;
       END_IF;
   END_FOR;
   "FRK_DecisionCyclic"(Owner := #Root,
                        Busy := FALSE,
                        Reset := TRUE,
                        AlarmLog := "GDB_DecisionTest".Log);
   "FRK_DecisionCyclic"(Owner := #Peer,
                        Busy := FALSE,
                        Reset := TRUE,
                        AlarmLog := "GDB_DecisionTest".Log);
   "GDB_DecisionTest".Done := TRUE;
END_FUNCTION

FUNCTION "F_TestEventSink" : Void   // FC1, SCL
{ S7_Optimized_Access := 'TRUE' }
VERSION : 0.1
// stored: AutoNumber true, IsIECCheckEnabled false, SetENOAutomatically false, UDAEnableTagReadback false
   VAR_INPUT
      Ev : "ST_AlarmEvent";
   END_VAR
BEGIN

   "GDB_StateAlarmTest".SinkLast := #Ev;
   IF #Ev.State = 0 THEN
       "GDB_StateAlarmTest".SinkClose := "GDB_StateAlarmTest".SinkClose + 1;
   ELSE
       "GDB_StateAlarmTest".SinkCome := "GDB_StateAlarmTest".SinkCome + 1;
   END_IF;
END_FUNCTION

DATA_BLOCK "GDB_FraktalMain"   // DB28
VERSION : 0.1
// stored: AutoNumber true, DBAccessibleFromOPCUA true, DBAccessibleFromWebserver true, InstanceOfName FB_FraktalMain, InstanceOfType FB
"FB_FraktalMain"
BEGIN
END_DATA_BLOCK

DATA_BLOCK "StationA"   // DB25
VERSION : 0.1
// stored: AutoNumber true, DBAccessibleFromOPCUA true, DBAccessibleFromWebserver true, InstanceOfName FB_DeclarationUnit, InstanceOfType FB
"FB_DeclarationUnit"
BEGIN
END_DATA_BLOCK

DATA_BLOCK "StationB"   // DB26
VERSION : 0.1
// stored: AutoNumber true, DBAccessibleFromOPCUA true, DBAccessibleFromWebserver true, InstanceOfName FB_DeclarationUnit, InstanceOfType FB
"FB_DeclarationUnit"
BEGIN
END_DATA_BLOCK
